# EPICS autosave request: iocs/meascomp/db/measCompAnalogOut_settings.req
$(P)$(R)Pulse
$(P)$(R)Range
$(P)$(R)TweakVal
$(P)$(R).DRVL
$(P)$(R).DRVH
$(P)$(R).LOPR
$(P)$(R).HOPR
$(P)$(R).EGUF
$(P)$(R).EGUL
$(P)$(R).PREC
$(P)$(R)Return.DRVL
$(P)$(R)Return.DRVH
$(P)$(R)Return.LOPR
$(P)$(R)Return.HOPR
$(P)$(R)Return.EGUF
$(P)$(R)Return.EGUL
$(P)$(R)Return.PREC
$(P)$(R)SyncMaster
$(P)$(R)SyncEnable
